Yaskawa INFORM job: ENDDETPRG.JBI

/JOB
//NAME ENDDETPRG
///FOLDERNAME FOLDER003
//POS
///NPOS 0,0,0,0,0,0
//INST
///DATE 2017/04/26 10:21
///ATTR SC,RW
///GROUP1 RB1
NOP
SKILLSND "ENDDET"
ADVINIT
END
